SUBAPPLICATION Uebung_094b4b_AX (* Wie Uebung_094b_AX, aber mit MyLib::sys::NumericValue_TO_AUI2_AND_STORE als wiederverwendbarem Baustein: wie NumericValue_TO_AUI2 (bidirektionaler VALUEO-Plug direkt an AOption_AUI_DEMUX_2.K), zusaetzlich mit INI-Persistenz des Index. *)
  (* Standard: 61499-2; Description: Copyright (c) 2026 Meisterschulen am Ostbahnhof This program and the accompanying materials are made available under the terms of the Eclipse Public License 2.0 which is available at https://www.eclipse.org/legal/epl-2.0/ SPDX-License-Identifier: EPL-2.0 *)
  (* Version 1.1, 2026-10-13, Franz Höpfinger, Meisterschulen am Ostbahnhof, NumericValue_TO_AUI2 ersetzt durch NumericValue_TO_AUI2_AND_STORE - gleicher bidirektionaler VALUEO-Plug, zusaetzlich INI-persistiert (KEY_I1_STORE/SECTION_I1_STORE, bereits aus Uebung_012c_AUDI bekannt). *)
  PACKAGE Uebungen;
  IMPORT Uebungen::const::NVS::NVS_Keys::KEY_I1_STORE;
  IMPORT Uebungen::const::NVS::NVS_Keys::SECTION_I1_STORE;
  IMPORT Uebungen::const::UT::DefaultPool::InputNumber_I1;
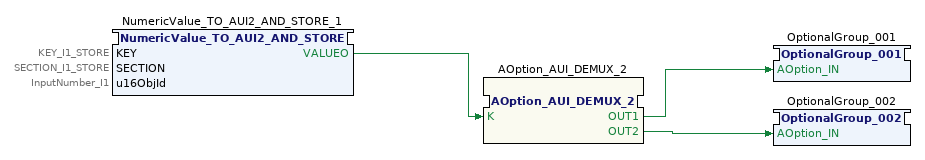
  FBS
    AOption_AUI_DEMUX_2 : Option::selection::AOption_AUI_DEMUX_2;
  END_FBS
  SUBAPPS
    NumericValue_TO_AUI2_AND_STORE_1 : MyLib::sys::NumericValue_TO_AUI2_AND_STORE(KEY := KEY_I1_STORE, SECTION := SECTION_I1_STORE, u16ObjId := InputNumber_I1);
    OptionalGroup_001 : MyLib_AX_Option::sys::OptionalGroup_001;
    OptionalGroup_002 : MyLib_AX_Option::sys::OptionalGroup_002;
  END_SUBAPPS
  ADAPTER_CONNECTIONS
    NumericValue_TO_AUI2_AND_STORE_1.VALUEO TO AOption_AUI_DEMUX_2.K;
    AOption_AUI_DEMUX_2.OUT1 TO OptionalGroup_001.AOption_IN;
    AOption_AUI_DEMUX_2.OUT2 TO OptionalGroup_002.AOption_IN;
  END_CONNECTIONS
END_SUBAPPLICATION
